(* IEC 61131-3 sources: ecmccfg/examples/PSI/lab_setup/block_motion_funcs/cfg, 3 files *)

(* ---- block_motion_funcs.plc ---- *)
# Block ordinary motion during an interlock-controlled parking home.
#
# Test operation:
#   1. Set this PLC's debug input high to assert the test interlock.
#   2. The PLC blocks ABS/REL/velocity commands, stops existing motion and
#      starts homing procedure 1. Homing remains admitted.
#   3. While homing, send arbitrary motor-record or native ABS commands. They
#      must be ignored without changing the active homing execute state.
#   4. Native/motor STOP and disable commands remain effective by design.
#
# Cfg.SetAxisIgnoreDisabledMotionCommands(AID,1) is configured permanently in
# startup.cmd. Do not toggle that policy here: when all motion functions are
# enabled it has no effect, and keeping it enabled closes transition races.

VAR
  AID                     : 1;
  HOME_SEQUENCE           : 1;
  HOME_VEL_TO             : 4;
  HOME_VEL_FROM           : 0.5;
  HOME_POSITION           : -55;
  HOME_TIMEOUT_SEC        : 30;

  ax_enabled              : ax1.drv.enabled;

  state                   : static.state;
  interlock               : static.interlock;
  interlock_old           : static.interlock_old;
  home_started            : static.home_started;
  timeout_cycles          : static.timeout_cycles;

  FALSE                   : 0;
  TRUE                    : 1;
  NOT_BUSY                : 0;
  BUSY                    : 1;

  SM_BOOT                 : 0;
  SM_IDLE                 : 10;
  SM_STOP                 : 20;
  SM_ENABLE               : 30;
  SM_START_HOME           : 40;
  SM_WAIT_HOME            : 50;
  SM_DISABLE              : 60;
END_VAR

if(${SELF}.firstscan) {
  state := SM_BOOT;
  interlock := FALSE;
  interlock_old := FALSE;
  home_started := FALSE;
  timeout_cycles := 0;
};

# The PLC debug input is the reproducible test-interlock source.
if(state != SM_BOOT) {
  if(${SELF}.dbg == TRUE) {
    interlock := TRUE;
  }
  else {
    interlock := FALSE;
  };
};

if(state == SM_BOOT) {
  if(epics_get_started() == TRUE) {
    mc_set_enable_motion_funcs(AID, 1, 1, 1);
    state := SM_IDLE;
    println('block_motion_funcs: ready');
  };
}

else if(state == SM_IDLE) {
  if((interlock == TRUE) and (interlock_old == FALSE)) {
    # Close command admission before touching the active trajectory. ABS/REL,
    # PVT and velocity/jog requests are now ignored, while HOME stays allowed.
    mc_set_enable_motion_funcs(AID, 0, 0, 1);
    home_started := FALSE;

    # Use the native synchronous command path. Motor-record STOP/CNEN requests
    # are asynchronous and can otherwise arrive after a new home has started.
    # Native disable is intentionally not filtered by the motion-function gate.
    mc_power(AID, 0);
    state := SM_STOP;
    println('block_motion_funcs: moves blocked; disabling active motion');
  }
  else if(interlock == FALSE) {
    # Ignore mode remains configured, but no command type is disabled here.
    mc_set_enable_motion_funcs(AID, 1, 1, 1);
  };
}

else if(state == SM_STOP) {
  # Do not start home until both trajectory and drive acknowledge the native
  # disable. This prevents a late disable from cancelling the new home.
  if((mc_get_busy(AID) == NOT_BUSY) and (ax_enabled == FALSE)) {
    state := SM_ENABLE;
  };
}

else if(state == SM_ENABLE) {
  if(ax_enabled == FALSE) {
    mc_power(AID, 1);
  }
  else {
    state := SM_START_HOME;
  };
}

else if(state == SM_START_HOME) {
  # Generate one explicit low-to-high home edge.
  mc_home_pos(AID, 0, HOME_SEQUENCE,
              HOME_VEL_TO, HOME_VEL_FROM, HOME_POSITION);
  mc_home_pos(AID, 1, HOME_SEQUENCE,
              HOME_VEL_TO, HOME_VEL_FROM, HOME_POSITION);
  timeout_cycles := HOME_TIMEOUT_SEC / ${SELF}.scantime;
  state := SM_WAIT_HOME;
  println('block_motion_funcs: homing requested');
}

else if(state == SM_WAIT_HOME) {
  timeout_cycles := timeout_cycles - 1;

  # Require observation of an active home. This prevents an old Homed=1 value
  # from completing the state before the new request has actually run.
  if(mc_get_busy(AID) == BUSY) {
    home_started := TRUE;
  };

  if((home_started == TRUE)
     and (mc_get_busy(AID) == NOT_BUSY)
     and (mc_get_homed(AID) == TRUE)) {
    state := SM_DISABLE;
    println('block_motion_funcs: homing complete');
  }
  else if((home_started == TRUE)
          and (mc_get_busy(AID) == NOT_BUSY)
          and (mc_get_homed(AID) == FALSE)) {
    # An external native/motor STOP or disable must remain effective. Treat it
    # as an aborted home and finish in the safe disabled state.
    state := SM_DISABLE;
    println('block_motion_funcs: homing aborted by STOP or disable');
  }
  else if(timeout_cycles < 0) {
    state := SM_DISABLE;
    println('block_motion_funcs: homing timeout');
  };
}

else if(state == SM_DISABLE) {
  # Native disable is deliberate and must remain effective even while ordinary
  # motion functions are blocked.
  mc_power(AID, 0);

  if(ax_enabled == FALSE) {
    home_started := FALSE;
    state := SM_IDLE;

    if(interlock == FALSE) {
      mc_set_enable_motion_funcs(AID, 1, 1, 1);
    };
    println('block_motion_funcs: parked and disabled');
  };
};

interlock_old := interlock;
# vim: set expandtab ts=2 sw=2 sts=2 et:

(* ---- test.plc ---- *)
#
# file:   eht_interlock_parking.plc
# author: Felix Maier <felix.maier@psi.ch>, November 2026
#
# This PLC code moves the EHT "lifting X" axis to the parking position when an
# interlock is detected. The default park position is the right side (looking
# in beam direction).  # This can be changed by setting the PV
# `PREFIX:X-ParkPos' to LEFT.  Configuration for speed, acceleration, timeout
# and the actual parking positions in mm can be configured in the below VAR
# section.
#
# TODO:
#   - only one parking position is possible, due to homing.
#   - mc_set_enable_motion_funcs: connect it to the flag is_pending_interlock.
#   - add PV with interlock flag.

VAR
  # configuration
  AID                     :   1;
  PARK_VEL                :   3;
  PARK_VEL_SLOW           :   0.5;
  PARK_ACC                :   2;
  PARK_POS_LEFT_MM        :   60;
  PARK_POS_RIGHT_MM       :   5.3;
  TIMEOUT_SEC             :   20;

  # pv
  pv_park_position        :   static.pv_park_position;

  prev_dbg                :   static.prev_dbg;

  # axis
  ax_enabled              :   ax1.drv.enabled;
  ax_actpos               :   ax1.enc.actpos;

  # variables
  prev_is_interlock       :   static.prev_is_interlock;
  prev_pv_park_position   :   static.prev_park_position;
  timeout_cycles          :   static.timeout_cycles;
  is_interlock            :   static.is_interlock;
  is_pend_interlock       :   static.is_pend_interlock;
  park_position           :   static.park_position;

  # constants
  TRUE                    :   1;
  FALSE                   :   0;
  BUSY                    :   1;
  NOT_BUSY                :   0;
  PV_PARK_RIGHT           :   0;
  PV_PARK_LEFT            :   1;
  PARK_TOL                :   0.5;

  # error
  ERROR_TIMEOUT           :   262144; # 0x40000

  # state machine
  state                   :   static.state;
  SM_BOOT                 :   2;
  SM_IDLE                 :   0;
  SM_INIT                 :   100;
  SM_START_MOVE           :   200;
  SM_START_MOVE2          :   250;
  SM_WAIT_FOR_PARKING     :   300;
  SM_DISABLE              :   400;

END_VAR

# -----------------------------------------------------------------------------
if(${SELF}.firstscan) {
  state := SM_BOOT;
  timeout_cycles := TIMEOUT_SEC / ${SELF}.scantime;
  park_position := PARK_POS_RIGHT_MM;
  is_pend_interlock := FALSE;
  is_interlock := FALSE;
};

# =============================================================================
# INTERLOCK & TIMEOUT HANDLING
# =============================================================================
if(state != SM_BOOT) {
  if(${SELF}.dbg  == TRUE) {
    is_interlock := TRUE;
  }
  else {
    is_interlock := FALSE;
  };

  if (state != SM_IDLE) {
    timeout_cycles := timeout_cycles - 1;

    if (timeout_cycles < 0) {
      #mc_set_axis_error(AID, ERROR_TIMEOUT);
      #state := SM_DISABLE;
    };
  }
}

# =============================================================================
# STATES
# =============================================================================
if (state == SM_BOOT) {
  if(epics_get_started() == TRUE) {
    state := SM_IDLE;
  }
}

else if (state == SM_IDLE) {
  if( (is_interlock == TRUE) and (prev_is_interlock == FALSE) ) {
    println('__EHT__: interlock detected');
    if(mc_get_busy(AID) == BUSY) {

      println('__EHT__: axis is moving, halt');
      mc_mr_set_cnen(AID, 0);
      mc_mr_set_stop(AID, 1);
    };
    is_pend_interlock := TRUE;
    state := SM_INIT;
    println('__EHT__: state -> SM_INIT');
    println('__EHT__: disable motion functions');
    mc_set_enable_motion_funcs(AID, 0, 0, 1);
    mc_set_ignore_disabled_motion_cmds(AID,1);
    timeout_cycles := TIMEOUT_SEC / ${SELF}.scantime;
  }
  else if( (is_interlock == FALSE) and (prev_is_interlock == TRUE) ) {
    println('__EHT__: enable move functions');
    is_pend_interlock := FALSE;
    mc_set_enable_motion_funcs(AID, 1, 1, 1);
    mc_set_ignore_disabled_motion_cmds(AID,0);
  }

  if( (is_pend_interlock == TRUE) and (ax_enabled) ) {
    mc_mr_set_cnen(AID, 0);
  }

  # change park position
  if( (prev_pv_park_position == PV_PARK_RIGHT) and (pv_park_position == PV_PARK_LEFT) ) {
    println('__EHT__: change park position to LEFT');
    park_position := PARK_POS_LEFT_MM;
  };

  if( (prev_pv_park_position == PV_PARK_LEFT) and (pv_park_position == PV_PARK_RIGHT) ) {
    println('__EHT__: change park position to Right');
    park_position := PARK_POS_RIGHT_MM;
  };
}

else if (state == SM_INIT) {
  if(mc_get_busy(AID) == NOT_BUSY) {
    if( ax_enabled == TRUE) {
      state := SM_START_MOVE;
      println('__EHT__: state -> SM_START_MOVE');
    }
    else {
      mc_power(AID, 1);
    };
  };
}

else if (state == SM_START_MOVE) {
  mc_home_pos(AID, 0, 1, PARK_VEL, PARK_VEL_SLOW, -55);
  mc_home_pos(AID, 1, 1, PARK_VEL, PARK_VEL_SLOW, -55);
  println('__EHT__: ---------------------------> DEBUG');
  if(mc_get_busy(AID) == BUSY) {
    state := SM_WAIT_FOR_PARKING;
    println('__EHT__: state -> SM_WAIT_FOR_PARKING');
  }
}

else if (state == SM_WAIT_FOR_PARKING) {
  if(mc_get_homed(AID)) {
    state := SM_DISABLE;
    println('__EHT__: state -> SM_DISABLE');
  };
}

else if (state == SM_DISABLE) {
  #mc_power(AID,0);
  mc_mr_set_cnen(AID, 0);
  state := SM_IDLE;
  if(is_interlock == FALSE) {
    println('__EHT__: enable move functions');
    mc_set_enable_motion_funcs(AID, 1, 1, 1);
    mc_set_ignore_disabled_motion_cmds(AID,0);
  }
  println('__EHT__: state -> SM_IDLE');
};

# -----------------------------------------------------------------------------
prev_dbg := ${SELF}.dbg;
prev_is_interlock := is_interlock;
prev_pv_park_position := pv_park_position;
# vim: set expandtab ts=2 sw=2 sts=2 et:

(* ---- test_slimmed_down.plc ---- *)
VAR
  AID                     :   1;

  ax_enabled              :   ax1.drv.enabled;
  prev_is_interlock       :   static.prev_is_interlock;
  is_interlock            :   static.is_interlock;
  is_pend_interlock       :   static.is_pend_interlock;

  # constants
  TRUE                    :   1;
  FALSE                   :   0;
  BUSY                    :   1;
  NOT_BUSY                :   0;

  # state machine
  state                   :   static.state;
  SM_BOOT                 :   2;
  SM_IDLE                 :   0;
  SM_INIT                 :   100;
  SM_START_MOVE           :   200;
  SM_START_MOVE2          :   250;
  SM_WAIT_FOR_PARKING     :   300;
  SM_DISABLE              :   400;

END_VAR

# -----------------------------------------------------------------------------
if(${SELF}.firstscan) {
  state := SM_BOOT;
  is_pend_interlock := FALSE;
  is_interlock := FALSE;
};

if(state != SM_BOOT) {
  if(${SELF}.dbg  == TRUE) {
    is_interlock := TRUE;
  }
  else {
    is_interlock := FALSE;
  };
}

# =============================================================================
# STATES
# =============================================================================
if (state == SM_BOOT) {
  if(epics_get_started() == TRUE) {
    state := SM_IDLE;
  }
}

else if (state == SM_IDLE) {
  if( (is_interlock == TRUE) and (prev_is_interlock == FALSE) ) {
    if(mc_get_busy(AID) == BUSY) {
      println('__EHT__: axis is moving, halt');
      mc_power(AID, 0);
      #mc_mr_set_cnen(AID, 0);
      #mc_mr_set_stop(AID, 1);
    };
    is_pend_interlock := TRUE;
    state := SM_INIT;
    mc_set_enable_motion_funcs(AID, 0, 0, 1);
    mc_set_ignore_disabled_motion_cmds(AID,1);
  }
  else if( (is_interlock == FALSE) and (prev_is_interlock == TRUE) ) {
    is_pend_interlock := FALSE;
    mc_set_enable_motion_funcs(AID, 1, 1, 1);
    mc_set_ignore_disabled_motion_cmds(AID,0);
  }

  if( (is_pend_interlock == TRUE) and (ax_enabled) ) {
    mc_mr_set_cnen(AID, 0);
  }
}

else if (state == SM_INIT) {
  if(mc_get_busy(AID) == NOT_BUSY) {
    if( ax_enabled == TRUE) {
      state := SM_START_MOVE;
    }
    else {
      mc_power(AID, 1);
    };
  };
}

else if (state == SM_START_MOVE) {
  mc_home_pos(AID, 0, 1, 4, 0.5, -55);
  mc_home_pos(AID, 1, 1, 4, 0.5, -55);
  state := SM_WAIT_FOR_PARKING;
}

else if (state == SM_WAIT_FOR_PARKING) {
  if(mc_get_homed(AID)) {
    state := SM_DISABLE;
  };
}

else if (state == SM_DISABLE) {
  mc_mr_set_cnen(AID, 0);
  state := SM_IDLE;
  if(is_interlock == FALSE) {
    mc_set_enable_motion_funcs(AID, 1, 1, 1);
    mc_set_ignore_disabled_motion_cmds(AID,0);
  }
};

# -----------------------------------------------------------------------------

prev_is_interlock := is_interlock;
# vim: set expandtab ts=2 sw=2 sts=2 et:
